(* IEC 61131-3 sources: volt/packages/volt-lsp-iec/test-corpus/awa-palletizer/Device/Plc Logic/Application/Library Manager/(unresolved)/cmpusermgr implementation, 51 files *)

(* ---- USERMGRCHANGEMYPASSWORD.pou ---- *)
FUNCTION USERMGRCHANGEMYPASSWORD : RTS_IEC_RESULT
VAR_INPUT
	HUSER : RTS_IEC_HANDLE;
	PSZUSER : REFERENCE TO STRING;
	PSZOLDPASSWORD : REFERENCE TO STRING;
	PSZNEWPASSWORD : REFERENCE TO STRING;
END_VAR
END_FUNCTION

(* ---- USERMGRGETSESSIONUSER.pou ---- *)
FUNCTION USERMGRGETSESSIONUSER : RTS_IEC_HANDLE
VAR_INPUT
	SESSIONID : UDINT;
	PRESULT : POINTER TO RTS_IEC_RESULT;
END_VAR
END_FUNCTION

(* ---- USERMGRGETUSERACCESSRIGHTS.pou ---- *)
FUNCTION USERMGRGETUSERACCESSRIGHTS : RTS_IEC_RESULT
VAR_INPUT
	PSZOBJECT : REFERENCE TO STRING;
	HUSER : RTS_IEC_HANDLE;
	PULRIGHTS : POINTER TO DWORD;
	PULDENIEDRIGHTS : POINTER TO DWORD;
END_VAR
END_FUNCTION

(* ---- USERMGRGROUPADD.pou ---- *)
FUNCTION USERMGRGROUPADD : RTS_IEC_RESULT
VAR_INPUT
	HUSER : RTS_IEC_HANDLE;
END_VAR
VAR_IN_OUT
	PSZGROUPNAME : STRING;
END_VAR
END_FUNCTION

(* ---- USERMGRGROUPADDUSER.pou ---- *)
FUNCTION USERMGRGROUPADDUSER : RTS_IEC_RESULT
VAR_INPUT
	HUSER : RTS_IEC_HANDLE;
END_VAR
VAR_IN_OUT
	PSZGROUPNAME : STRING;
	PSZUSERNAME : STRING;
END_VAR
END_FUNCTION

(* ---- USERMGRGROUPGETFIRST.pou ---- *)
FUNCTION USERMGRGROUPGETFIRST : RTS_IEC_HANDLE
VAR_INPUT
	HUSER : RTS_IEC_HANDLE;
END_VAR
VAR_OUTPUT
	RESULT : RTS_IEC_RESULT;
END_VAR
END_FUNCTION

(* ---- USERMGRGROUPGETFIRSTUSER.pou ---- *)
FUNCTION USERMGRGROUPGETFIRSTUSER : RTS_IEC_RESULT
VAR_INPUT
	HUSER : RTS_IEC_HANDLE;
	HGROUP : RTS_IEC_HANDLE;
END_VAR
VAR_IN_OUT
	PHITERATOR : RTS_IEC_HANDLE;
	PSZUSERNAME : STRING(59);
END_VAR
END_FUNCTION

(* ---- USERMGRGROUPGETFIRSTUSERINTERNAL.pou ---- *)
FUNCTION USERMGRGROUPGETFIRSTUSERINTERNAL : RTS_IEC_RESULT
VAR_INPUT
	HUSER : RTS_IEC_HANDLE;
	HGROUP : RTS_IEC_HANDLE;
	IMAXLEN : UDINT;
END_VAR
VAR_IN_OUT
	PHITERATOR : RTS_IEC_HANDLE;
	PSZUSERNAME : STRING;
END_VAR
END_FUNCTION

(* ---- USERMGRGROUPGETHANDLE.pou ---- *)
FUNCTION USERMGRGROUPGETHANDLE : RTS_IEC_HANDLE
VAR_INPUT
	HUSER : RTS_IEC_HANDLE;
END_VAR
VAR_OUTPUT
	RESULT : RTS_IEC_RESULT;
END_VAR
VAR_IN_OUT
	PSZGROUPNAME : STRING;
END_VAR
END_FUNCTION

(* ---- USERMGRGROUPGETNAME.pou ---- *)
FUNCTION USERMGRGROUPGETNAME : RTS_IEC_RESULT
VAR_INPUT
	HUSER : RTS_IEC_HANDLE;
	HGROUP : RTS_IEC_HANDLE;
END_VAR
VAR_IN_OUT
	PSZGROUP : STRING(59);
END_VAR
END_FUNCTION

(* ---- USERMGRGROUPGETNAMEINTERNAL.pou ---- *)
FUNCTION USERMGRGROUPGETNAMEINTERNAL : RTS_IEC_RESULT
VAR_INPUT
	HUSER : RTS_IEC_HANDLE;
	HGROUP : RTS_IEC_HANDLE;
	IMAXLEN : UDINT;
END_VAR
VAR_IN_OUT
	PSZGROUP : STRING;
END_VAR
END_FUNCTION

(* ---- USERMGRGROUPGETNEXT.pou ---- *)
FUNCTION USERMGRGROUPGETNEXT : RTS_IEC_HANDLE
VAR_INPUT
	HUSER : RTS_IEC_HANDLE;
	HPREVGROUP : RTS_IEC_HANDLE;
END_VAR
VAR_OUTPUT
	RESULT : RTS_IEC_RESULT;
END_VAR
END_FUNCTION

(* ---- USERMGRGROUPGETNEXTUSER.pou ---- *)
FUNCTION USERMGRGROUPGETNEXTUSER : RTS_IEC_RESULT
VAR_INPUT
	HUSER : RTS_IEC_HANDLE;
	HGROUP : RTS_IEC_HANDLE;
END_VAR
VAR_IN_OUT
	PHITERATOR : RTS_IEC_HANDLE;
	PSZUSERNAME : STRING(59);
END_VAR
END_FUNCTION

(* ---- USERMGRGROUPGETNEXTUSERINTERNAL.pou ---- *)
FUNCTION USERMGRGROUPGETNEXTUSERINTERNAL : RTS_IEC_RESULT
VAR_INPUT
	HUSER : RTS_IEC_HANDLE;
	HGROUP : RTS_IEC_HANDLE;
	IMAXLEN : UDINT;
END_VAR
VAR_IN_OUT
	PHITERATOR : RTS_IEC_HANDLE;
	PSZUSERNAME : STRING;
END_VAR
END_FUNCTION

(* ---- USERMGRGROUPREMOVE.pou ---- *)
FUNCTION USERMGRGROUPREMOVE : RTS_IEC_RESULT
VAR_INPUT
	HUSER : RTS_IEC_HANDLE;
END_VAR
VAR_IN_OUT
	PSZGROUPNAME : STRING;
END_VAR
END_FUNCTION

(* ---- USERMGRGROUPREMOVEUSER.pou ---- *)
FUNCTION USERMGRGROUPREMOVEUSER : RTS_IEC_RESULT
VAR_INPUT
	HUSER : RTS_IEC_HANDLE;
END_VAR
VAR_IN_OUT
	PSZGROUP : STRING;
	PSZUSER : STRING;
END_VAR
END_FUNCTION

(* ---- USERMGRHASUSERACCESSRIGHTS.pou ---- *)
FUNCTION USERMGRHASUSERACCESSRIGHTS : RTS_IEC_RESULT
VAR_INPUT
	PSZOBJECT : REFERENCE TO STRING;
	HUSER : RTS_IEC_HANDLE;
	ULREQUESTEDRIGHTS : DWORD;
END_VAR
END_FUNCTION

(* ---- USERMGRISACTIVE.pou ---- *)
FUNCTION USERMGRISACTIVE : BOOL
END_FUNCTION

(* ---- USERMGRLOGIN.pou ---- *)
FUNCTION USERMGRLOGIN : RTS_IEC_HANDLE
VAR_INPUT
	PSZUSER : REFERENCE TO STRING;
	PSZPASSWORD : REFERENCE TO STRING;
	PRESULT : POINTER TO RTS_IEC_RESULT;
END_VAR
END_FUNCTION

(* ---- USERMGRLOGOUT.pou ---- *)
FUNCTION USERMGRLOGOUT : RTS_IEC_RESULT
VAR_INPUT
	HUSER : RTS_IEC_HANDLE;
END_VAR
END_FUNCTION

(* ---- USERMGROBJECTADD.pou ---- *)
FUNCTION USERMGROBJECTADD : RTS_IEC_HANDLE
VAR_INPUT
	PSZOBJECT : REFERENCE TO STRING;
	PRESULT : POINTER TO RTS_IEC_RESULT;
END_VAR
END_FUNCTION

(* ---- USERMGROBJECTADDGROUP.pou ---- *)
FUNCTION USERMGROBJECTADDGROUP : RTS_IEC_RESULT
VAR_INPUT
	HUSER : RTS_IEC_HANDLE;
	HOBJECT : RTS_IEC_HANDLE;
	HGROUP : RTS_IEC_HANDLE;
END_VAR
END_FUNCTION

(* ---- USERMGROBJECTCLEARRIGHTS.pou ---- *)
FUNCTION USERMGROBJECTCLEARRIGHTS : RTS_IEC_RESULT
VAR_INPUT
	HUSER : RTS_IEC_HANDLE;
	HOBJECT : RTS_IEC_HANDLE;
END_VAR
END_FUNCTION

(* ---- USERMGROBJECTGETFIRSTCHILD.pou ---- *)
FUNCTION USERMGROBJECTGETFIRSTCHILD : RTS_IEC_HANDLE
VAR_INPUT
	HFATHEROBJECT : RTS_IEC_HANDLE;
END_VAR
VAR_OUTPUT
	RESULT : RTS_IEC_RESULT;
END_VAR
END_FUNCTION

(* ---- USERMGROBJECTGETFIRSTGROUP.pou ---- *)
FUNCTION USERMGROBJECTGETFIRSTGROUP : RTS_IEC_HANDLE
VAR_INPUT
	HUSER : RTS_IEC_HANDLE;
	HOBJECT : RTS_IEC_HANDLE;
END_VAR
VAR_OUTPUT
	RESULT : RTS_IEC_RESULT;
END_VAR
END_FUNCTION

(* ---- USERMGROBJECTGETGROUPRIGHTS.pou ---- *)
FUNCTION USERMGROBJECTGETGROUPRIGHTS : RTS_IEC_RESULT
VAR_INPUT
	HUSER : RTS_IEC_HANDLE;
	HOBJECT : RTS_IEC_HANDLE;
	HGROUP : RTS_IEC_HANDLE;
END_VAR
VAR_OUTPUT
	ULRIGHTS : DWORD;
	ULDENIEDRIGHTS : DWORD;
END_VAR
END_FUNCTION

(* ---- USERMGROBJECTGETHANDLE.pou ---- *)
FUNCTION USERMGROBJECTGETHANDLE : RTS_IEC_HANDLE
VAR_OUTPUT
	RESULT : RTS_IEC_RESULT;
END_VAR
VAR_IN_OUT
	PSZOBJECTNAME : STRING;
END_VAR
END_FUNCTION

(* ---- USERMGROBJECTGETNAME.pou ---- *)
FUNCTION USERMGROBJECTGETNAME : RTS_IEC_RESULT
VAR_INPUT
	HOBJECT : RTS_IEC_HANDLE;
	PSZOBJECT : POINTER TO STRING;
	PIMAXLEN : POINTER TO UDINT;
END_VAR
END_FUNCTION

(* ---- USERMGROBJECTGETNEXTCHILD.pou ---- *)
FUNCTION USERMGROBJECTGETNEXTCHILD : RTS_IEC_HANDLE
VAR_INPUT
	HFATHEROBJECT : RTS_IEC_HANDLE;
	HPREVCHILD : RTS_IEC_HANDLE;
END_VAR
VAR_OUTPUT
	RESULT : RTS_IEC_RESULT;
END_VAR
END_FUNCTION

(* ---- USERMGROBJECTGETNEXTGROUP.pou ---- *)
FUNCTION USERMGROBJECTGETNEXTGROUP : RTS_IEC_HANDLE
VAR_INPUT
	HUSER : RTS_IEC_HANDLE;
	HOBJECT : RTS_IEC_HANDLE;
	HPREVGROUP : RTS_IEC_HANDLE;
END_VAR
VAR_OUTPUT
	RESULT : RTS_IEC_RESULT;
END_VAR
END_FUNCTION

(* ---- USERMGROBJECTREMOVE.pou ---- *)
FUNCTION USERMGROBJECTREMOVE : RTS_IEC_RESULT
VAR_INPUT
	HOBJECT : RTS_IEC_HANDLE;
END_VAR
END_FUNCTION

(* ---- USERMGROBJECTREMOVEGROUP.pou ---- *)
FUNCTION USERMGROBJECTREMOVEGROUP : RTS_IEC_RESULT
VAR_INPUT
	HUSER : RTS_IEC_HANDLE;
	HOBJECT : RTS_IEC_HANDLE;
	HGROUP : RTS_IEC_HANDLE;
END_VAR
END_FUNCTION

(* ---- USERMGROBJECTSETGROUPDENIEDRIGHTS.pou ---- *)
FUNCTION USERMGROBJECTSETGROUPDENIEDRIGHTS : RTS_IEC_RESULT
VAR_INPUT
	HUSER : RTS_IEC_HANDLE;
	HOBJECT : RTS_IEC_HANDLE;
	HGROUP : RTS_IEC_HANDLE;
	ULDENIEDRIGHTS : DWORD;
END_VAR
END_FUNCTION

(* ---- USERMGROBJECTSETGROUPRIGHTS.pou ---- *)
FUNCTION USERMGROBJECTSETGROUPRIGHTS : RTS_IEC_RESULT
VAR_INPUT
	HUSER : RTS_IEC_HANDLE;
	HOBJECT : RTS_IEC_HANDLE;
	HGROUP : RTS_IEC_HANDLE;
	ULRIGHTS : DWORD;
END_VAR
END_FUNCTION

(* ---- USERMGROBJECTSETUSEDRIGHTS.pou ---- *)
FUNCTION USERMGROBJECTSETUSEDRIGHTS : RTS_IEC_RESULT
VAR_INPUT
	HOBJECT : RTS_IEC_HANDLE;
	ULUSEDRIGHTS : DWORD;
END_VAR
END_FUNCTION

(* ---- USERMGRRELOGIN.pou ---- *)
FUNCTION USERMGRRELOGIN : RTS_IEC_RESULT
VAR_INPUT
	HUSER : RTS_IEC_HANDLE;
	PSZUSER : REFERENCE TO STRING;
	PSZPASSWORD : REFERENCE TO STRING;
END_VAR
END_FUNCTION

(* ---- USERMGRUSERADD.pou ---- *)
FUNCTION USERMGRUSERADD : RTS_IEC_RESULT
VAR_INPUT
	HUSER : RTS_IEC_HANDLE;
END_VAR
VAR_IN_OUT
	PSZUSER : STRING;
	PCREDENTIALS : UserMgrCredentials;
END_VAR
END_FUNCTION

(* ---- USERMGRUSERADDINFOTOUSER.pou ---- *)
FUNCTION USERMGRUSERADDINFOTOUSER : RTS_IEC_RESULT
VAR_INPUT
	HUSER : RTS_IEC_HANDLE;
	KEY : __XWORD;
	VALUE : UserMgrCacheValue;
END_VAR
END_FUNCTION

(* ---- USERMGRUSERGETFIRST.pou ---- *)
FUNCTION USERMGRUSERGETFIRST : RTS_IEC_RESULT
VAR_INPUT
	HUSER : RTS_IEC_HANDLE;
END_VAR
VAR_OUTPUT
	USERPROPERTY : DWORD;
END_VAR
VAR_IN_OUT
	PHITERATOR : RTS_IEC_HANDLE;
	PSZUSERNAME : STRING(59);
END_VAR
END_FUNCTION

(* ---- USERMGRUSERGETFIRSTINTERNAL.pou ---- *)
FUNCTION USERMGRUSERGETFIRSTINTERNAL : RTS_IEC_RESULT
VAR_INPUT
	HUSER : RTS_IEC_HANDLE;
	IMAXLEN : UDINT;
END_VAR
VAR_OUTPUT
	USERPROPERTY : DWORD;
END_VAR
VAR_IN_OUT
	PHITERATOR : RTS_IEC_HANDLE;
	PSZUSERNAME : STRING;
END_VAR
END_FUNCTION

(* ---- USERMGRUSERGETINFOOFUSER.pou ---- *)
FUNCTION USERMGRUSERGETINFOOFUSER : DWORD
VAR_INPUT
	HUSER : RTS_IEC_HANDLE;
	KEY : __XWORD;
END_VAR
VAR_OUTPUT
	VALUE : UserMgrCacheValue;
END_VAR
END_FUNCTION

(* ---- USERMGRUSERGETNAME.pou ---- *)
FUNCTION USERMGRUSERGETNAME : RTS_IEC_RESULT
VAR_INPUT
	HUSER : RTS_IEC_HANDLE;
END_VAR
VAR_IN_OUT
	PSZUSERNAME : STRING(59);
END_VAR
END_FUNCTION

(* ---- USERMGRUSERGETNAMEINTERNAL.pou ---- *)
FUNCTION USERMGRUSERGETNAMEINTERNAL : RTS_IEC_RESULT
VAR_INPUT
	HUSER : RTS_IEC_HANDLE;
	IMAXLEN : UDINT;
END_VAR
VAR_IN_OUT
	PSZUSERNAME : STRING;
END_VAR
END_FUNCTION

(* ---- USERMGRUSERGETNEXT.pou ---- *)
FUNCTION USERMGRUSERGETNEXT : RTS_IEC_RESULT
VAR_INPUT
	HUSER : RTS_IEC_HANDLE;
END_VAR
VAR_OUTPUT
	USERPROPERTY : DWORD;
END_VAR
VAR_IN_OUT
	PHITERATOR : RTS_IEC_HANDLE;
	PSZUSERNAME : STRING(59);
END_VAR
END_FUNCTION

(* ---- USERMGRUSERGETNEXTINTERNAL.pou ---- *)
FUNCTION USERMGRUSERGETNEXTINTERNAL : RTS_IEC_RESULT
VAR_INPUT
	HUSER : RTS_IEC_HANDLE;
	IMAXLEN : UDINT;
END_VAR
VAR_OUTPUT
	USERPROPERTY : DWORD;
END_VAR
VAR_IN_OUT
	PHITERATOR : RTS_IEC_HANDLE;
	PSZUSERNAME : STRING;
END_VAR
END_FUNCTION

(* ---- USERMGRUSERGETPROPERTY.pou ---- *)
FUNCTION USERMGRUSERGETPROPERTY : DWORD
VAR_INPUT
	HUSER : RTS_IEC_HANDLE;
END_VAR
VAR_OUTPUT
	RESULT : RTS_IEC_RESULT;
END_VAR
VAR_IN_OUT
	PSZUSER : STRING;
END_VAR
END_FUNCTION

(* ---- USERMGRUSERREMOVE.pou ---- *)
FUNCTION USERMGRUSERREMOVE : RTS_IEC_RESULT
VAR_INPUT
	HUSER : RTS_IEC_HANDLE;
END_VAR
VAR_IN_OUT
	PSZUSER : STRING;
END_VAR
END_FUNCTION

(* ---- USERMGRUSERREMOVEINFOFROMALLUSERS.pou ---- *)
FUNCTION USERMGRUSERREMOVEINFOFROMALLUSERS : DWORD
VAR_INPUT
	KEY : __XWORD;
END_VAR
END_FUNCTION

(* ---- USERMGRUSERREMOVEINFOFROMUSER.pou ---- *)
FUNCTION USERMGRUSERREMOVEINFOFROMUSER : DWORD
VAR_INPUT
	HUSER : RTS_IEC_HANDLE;
	KEY : __XWORD;
END_VAR
END_FUNCTION

(* ---- USERMGRUSERSETCREDENTIALS.pou ---- *)
FUNCTION USERMGRUSERSETCREDENTIALS : RTS_IEC_RESULT
VAR_INPUT
	HUSER : RTS_IEC_HANDLE;
END_VAR
VAR_IN_OUT
	PSZUSER : STRING;
	PCREDENTIALS : UserMgrCredentials;
END_VAR
END_FUNCTION

(* ---- USERMGRUSERSETPROPERTY.pou ---- *)
FUNCTION USERMGRUSERSETPROPERTY : RTS_IEC_RESULT
VAR_INPUT
	HUSER : RTS_IEC_HANDLE;
	USERPROPERTY : DWORD;
END_VAR
VAR_IN_OUT
	PSZUSER : STRING;
END_VAR
END_FUNCTION
